ABB RAPID module: MAIN_1.prg

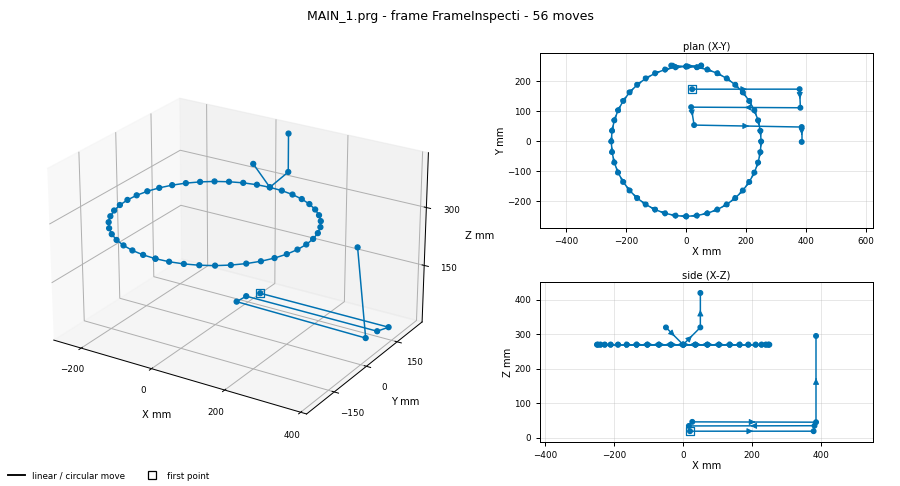
[picture p0: tool path of MAIN_1.prg in frame FrameInspecti, 56 of 76 moves have a stored position in this frame; points joined in program order, loops and branches not executed]
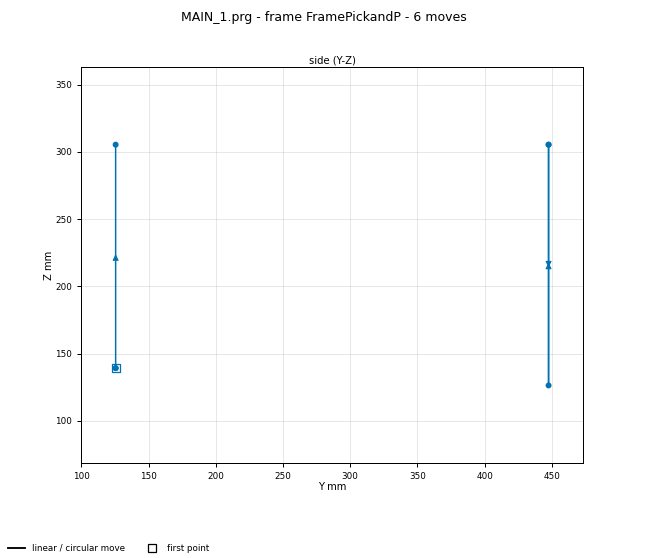
[picture p1: tool path of MAIN_1.prg in frame FramePickandP, 6 of 76 moves have a stored position in this frame; points joined in program order, loops and branches not executed]
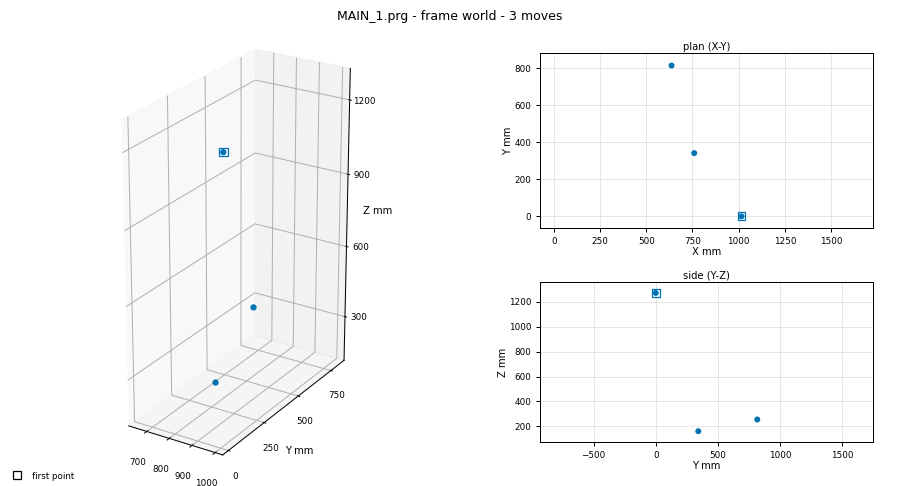
[picture p2: tool path of MAIN_1.prg in frame world, 3 of 76 moves have a stored position in this frame; points joined in program order, loops and branches not executed]
%%%
  VERSION:1
  LANGUAGE:ENGLISH
%%%
MODULE MOD_MAIN_1

    ! -------------------------------
    ! Define customized variables here
    ! ...

	! Tool variables:
	PERS tooldata Tool1 := [TRUE,[[129.073,0.000,85.477],[0.98018657,0.00000000,0.19807649,0.00000000]],[1,[0,0,20],[1,0,0,0],0,0,0.005]];
	PERS tooldata Tool1_withave := [TRUE,[[0.000,0.000,200.000],[1.00000000,0.00000000,0.00000000,0.00000000]],[1,[0,0,20],[1,0,0,0],0,0,0.005]];

	! Reference variables:
	PERS wobjdata FramePickandP := [FALSE, TRUE, "", [[719.013,-664.003,0.000],[1.00000000,0.00000000,0.00000000,0.00000000]],[[0,0,0],[1,0,0,0]]];
	PERS wobjdata FrameCircular := [FALSE, TRUE, "", [[577.670,392.250,0.000],[0.94275941,0.00000000,0.00000000,0.33347368]],[[0,0,0],[1,0,0,0]]];
	PERS wobjdata FrameInspecti := [FALSE, TRUE, "", [[0.000,782.714,377.610],[1.00000000,0.00000000,0.00000000,0.00000000]],[[0,0,0],[1,0,0,0]]];
	PERS wobjdata Frame1_withav := [FALSE, TRUE, "", [[0.000,1000.000,0.000],[1.00000000,0.00000000,0.00000000,0.00000000]],[[0,0,0],[1,0,0,0]]];

	PROC PROG1_withave()
		ConfJ \On;
		ConfL \Off;
		! This is a subprogram call to PROG_1
		MoveAbsJ [[-0.000001,0.000000,0.000000,0.000000,0.000000,-0.000000],[9E+09,9E+09,9E+09,9E+09,9E+09,9E+09]],v1000,z1,Tool1_withave \WObj:=Frame1_withav;
	ENDPROC

	PROC Main()
		ConfJ \On;
		ConfL \Off;
		! Program generated by RoboDK v5.6.9 for RoboDK Industrial on 26/02/2024 09:58:20
		! Using nominal kinematics.
		MoveAbsJ [[-0.000001,0.000000,0.000000,0.000000,0.000000,-0.000000],[9E+09,9E+09,9E+09,9E+09,9E+09,9E+09]],v500,z1,tool0 \WObj:=wobj0;
		MoveAbsJ [[0.000000,3.211240,-15.423700,0.000000,12.212500,-0.000000],[9E+09,9E+09,9E+09,9E+09,9E+09,9E+09]],v500,z1,tool0 \WObj:=wobj0;
		MoveL [[1015.000,0.000,1272.000],[0.70710678,0.00000000,0.70710678,0.00000001],[0,0,0,1],[9E+09,9E+09,9E+09,9E+09,9E+09,9E+09]],v500,z1,tool0 \WObj:=wobj0;
		SetDO D_OUT_5, 1;
		SetDO D_OUT_5, 1;
		SetDO D_OUT_5, 0.5;
		SetDO D_OUT_5, true;
		SetAO A_OUT_5, 1;
		SetAO A_OUT_5, 2;
		SetAO A_OUT_5, 0.5;
		SetAO A_OUT_5, true;
		SetDO var, val;
		SetAO var, val;
		WaitDI D_IN_5, 1;
		WaitDI D_IN_5, 1;
		WaitDI D_IN_5, 0.5;
		WaitDI D_IN_5, true;
		WaitDI D_IN_5, 1, \MaxTime:=0.1;
		WaitDI var, val;
		WaitDI var, val, \MaxTime:=0.1;
		TPWrite "Message";
		REMOTE_PROG_CALL_171;
		CODE_INSERT_172
		! Insert Comment
		MoveAbsJ [[-29.332200,46.677000,-0.024523,26.545600,25.395700,-51.634000],[9E+09,9E+09,9E+09,9E+09,9E+09,9E+09]],v500,z10,Tool1 \WObj:=FramePickandP;
		MoveL [[187.786,125.499,139.112],[0.00157079,-0.00002623,0.99999877,0.00003495],[-1,0,-1,0],[9E+09,9E+09,9E+09,9E+09,9E+09,9E+09]],v100,fine,Tool1 \WObj:=FramePickandP;
		SetDO D_OUT_5, 1;
		PICK_PART_111;
		MoveL CalcRobT([[-29.332200,46.677000,-0.024486,26.545800,25.395700,-51.634200],[9E+09,9E+09,9E+09,9E+09,9E+09,9E+09]],Tool1 \WObj:=FramePickandP),v300,z10,Tool1 \WObj:=FramePickandP;
		MoveL [[187.272,447.522,305.347],[0.00161443,0.00000875,0.99999870,-0.00001747],[-1,0,-1,0],[9E+09,9E+09,9E+09,9E+09,9E+09,9E+09]],v300,z10,Tool1 \WObj:=FramePickandP;
		! MoveSearch command not implemented
		MoveL [[187.851,447.517,126.235],[0.00161443,0.00000875,0.99999870,-0.00001747],[-1,0,-1,0],[9E+09,9E+09,9E+09,9E+09,9E+09,9E+09]],v100,fine,Tool1 \WObj:=FramePickandP;
		SetDO D_OUT_5, 0;
		PLACE_PART_112;
		MoveL [[187.272,447.522,305.347],[0.00161443,0.00000875,0.99999870,-0.00001747],[-1,0,-1,0],[9E+09,9E+09,9E+09,9E+09,9E+09,9E+09]],v100,z10,Tool1 \WObj:=FramePickandP;
		MoveAbsJ [[52.186000,45.675800,6.920000,66.734200,19.932300,-92.730000],[9E+09,9E+09,9E+09,9E+09,9E+09,9E+09]],v100,[FALSE,25.0,37.5,37.5,3.8,37.5,3.8],Tool1 \WObj:=FrameCircular;
		MoveC [[430.047,43.774,231.503],[0.08620627,-0.38531406,0.91758054,0.04634115],[0,0,-2,0],[9E+09,9E+09,9E+09,9E+09,9E+09,9E+09]],[[109.688,-153.222,161.073],[0.08620627,-0.38531406,0.91758054,0.04634115],[0,0,-2,0],[9E+09,9E+09,9E+09,9E+09,9E+09,9E+09]],v100,[FALSE,25.0,37.5,37.5,3.8,37.5,3.8],Tool1 \WObj:=FrameCircular;
		MoveC CalcRobT([[38.508400,52.810400,-4.822350,56.452300,29.788200,-93.025700],[9E+09,9E+09,9E+09,9E+09,9E+09,9E+09]], Tool1 \WObj:=FrameCircular),CalcRobT([[52.185900,45.675700,6.920040,66.734400,19.932300,-92.730300],[9E+09,9E+09,9E+09,9E+09,9E+09,9E+09]],Tool1 \WObj:=FrameCircular),v100,[FALSE,25.0,37.5,37.5,3.8,37.5,3.8],Tool1 \WObj:=FrameCircular;
		MoveL [[312.208,292.214,255.156],[0.08620627,-0.38531406,0.91758054,0.04634115],[0,0,-2,0],[9E+09,9E+09,9E+09,9E+09,9E+09,9E+09]],v100,fine,Tool1 \WObj:=FrameCircular;
		MoveAbsJ [[-0.000001,0.000000,0.000000,0.000000,0.000000,-0.000000],[9E+09,9E+09,9E+09,9E+09,9E+09,9E+09]],v100,fine,Tool1 \WObj:=FrameCircular;
		MoveAbsJ [[88.676000,29.601600,-6.428830,-1.984220,49.479200,4.547690],[9E+09,9E+09,9E+09,9E+09,9E+09,9E+09]],v100,fine,Tool1 \WObj:=FrameInspecti;
		MoveL [[19.898,174.307,19.008],[0.03212514,0.67543146,-0.73589088,0.03499889],[0,-1,0,0],[9E+09,9E+09,9E+09,9E+09,9E+09,9E+09]],v100,fine,Tool1 \WObj:=FrameInspecti;
		MoveL [[378.402,174.416,18.997],[0.03212514,0.67543146,-0.73589088,0.03499889],[0,0,-1,0],[9E+09,9E+09,9E+09,9E+09,9E+09,9E+09]],v100,fine,Tool1 \WObj:=FrameInspecti;
		MoveL [[380.996,112.363,34.882],[0.10687212,0.66688803,-0.72816340,0.11669088],[0,-1,-1,0],[9E+09,9E+09,9E+09,9E+09,9E+09,9E+09]],v100,fine,Tool1 \WObj:=FrameInspecti;
		MoveL [[16.551,114.359,34.226],[0.10687212,0.66688803,-0.72816340,0.11669088],[0,-1,0,0],[9E+09,9E+09,9E+09,9E+09,9E+09,9E+09]],v100,fine,Tool1 \WObj:=FrameInspecti;
		MoveL [[26.434,54.524,46.072],[0.02563823,-0.67223306,0.73935814,0.02819468],[0,-1,0,0],[9E+09,9E+09,9E+09,9E+09,9E+09,9E+09]],v100,fine,Tool1 \WObj:=FrameInspecti;
		MoveL [[385.448,48.050,45.137],[0.06581621,-0.66924184,0.73657112,0.07243323],[0,0,-1,0],[9E+09,9E+09,9E+09,9E+09,9E+09,9E+09]],v100,fine,Tool1 \WObj:=FrameInspecti;
		MoveL [[385.448,-1.625,295.251],[0.06581621,-0.66924184,0.73657112,0.07243323],[0,0,-1,0],[9E+09,9E+09,9E+09,9E+09,9E+09,9E+09]],v100,fine,Tool1 \WObj:=FrameInspecti;
		MoveAbsJ [[-0.000001,0.000000,0.000000,0.000000,0.000000,-0.000000],[9E+09,9E+09,9E+09,9E+09,9E+09,9E+09]],v100,fine,Tool1 \WObj:=FrameInspecti;
		EVENT_PROG_START_101;
		FrameInspecti := [FALSE, TRUE, "", [[13.637,-840.080,0.000],[0.70710678,0.00000000,0.00000000,-0.70710678]],[[0,0,0],[1,0,0,0]]];
		! Show Tool 1
		MoveAbsJ [[-68.090300,24.201900,26.785500,38.213400,36.201700,-98.796400],[9E+09,9E+09,9E+09,9E+09,9E+09,9E+09]],v1000,z1,Tool1 \WObj:=FrameInspecti;
		EVENT_PATH_APPROACH_102;
		MoveL [[-49.895,253.259,319.999],[0.00233251,-0.70710293,0.70710388,0.00202398],[-1,0,-2,0],[9E+09,9E+09,9E+09,9E+09,9E+09,9E+09]],v1000,z1,Tool1 \WObj:=FrameInspecti;
		MoveL [[0.000,250.000,270.000],[0.00233251,-0.70710293,0.70710388,0.00202398],[-1,0,-2,0],[9E+09,9E+09,9E+09,9E+09,9E+09,9E+09]],v1000,z1,Tool1 \WObj:=FrameInspecti;
		EVENT_PATH_START_103;
		MoveL [[35.579,247.455,270.000],[0.00259168,-0.70710203,0.70710482,0.00166608],[-1,0,-2,0],[9E+09,9E+09,9E+09,9E+09,9E+09,9E+09]],v50,z1,Tool1 \WObj:=FrameInspecti;
		MoveL [[70.433,239.873,270.000],[0.00280762,-0.70710738,0.70709946,0.00127734],[-1,0,-2,0],[9E+09,9E+09,9E+09,9E+09,9E+09,9E+09]],v50,z1,Tool1 \WObj:=FrameInspecti;
		MoveL [[103.854,227.408,270.000],[0.00295572,-0.70710677,0.70710008,0.00087007],[-1,0,-2,0],[9E+09,9E+09,9E+09,9E+09,9E+09,9E+09]],v50,z1,Tool1 \WObj:=FrameInspecti;
		MoveL [[135.160,210.313,270.000],[0.00305444,-0.70710635,0.70710047,0.00043812],[-1,0,-2,0],[9E+09,9E+09,9E+09,9E+09,9E+09,9E+09]],v50,z1,Tool1 \WObj:=FrameInspecti;
		MoveL [[163.715,188.937,270.000],[0.00308530,-0.70710622,0.70710061,0.00000001],[-1,0,-2,0],[9E+09,9E+09,9E+09,9E+09,9E+09,9E+09]],v50,z1,Tool1 \WObj:=FrameInspecti;
		MoveL [[188.937,163.715,270.000],[0.00305445,-0.70710635,0.70710047,-0.00043812],[-1,0,-2,0],[9E+09,9E+09,9E+09,9E+09,9E+09,9E+09]],v50,z1,Tool1 \WObj:=FrameInspecti;
		MoveL [[210.313,135.160,270.000],[0.00296806,-0.70710672,0.70710008,-0.00087007],[-1,0,-2,0],[9E+09,9E+09,9E+09,9E+09,9E+09,9E+09]],v50,z1,Tool1 \WObj:=FrameInspecti;
		MoveL [[227.408,103.854,270.000],[0.00281379,-0.70710735,0.70709945,-0.00128351],[-1,0,-2,0],[9E+09,9E+09,9E+09,9E+09,9E+09,9E+09]],v50,z1,Tool1 \WObj:=FrameInspecti;
		MoveL [[239.873,70.433,270.000],[0.00259785,-0.70710201,0.70710480,-0.00167225],[-1,0,-2,0],[9E+09,9E+09,9E+09,9E+09,9E+09,9E+09]],v50,z1,Tool1 \WObj:=FrameInspecti;
		MoveL [[247.455,35.579,270.000],[0.00233251,-0.70710293,0.70710388,-0.00202398],[-1,0,-2,0],[9E+09,9E+09,9E+09,9E+09,9E+09,9E+09]],v50,z1,Tool1 \WObj:=FrameInspecti;
		MoveL [[250.000,0.000,270.000],[0.00202398,-0.70710388,0.70710293,-0.00233251],[-1,0,-2,0],[9E+09,9E+09,9E+09,9E+09,9E+09,9E+09]],v50,z1,Tool1 \WObj:=FrameInspecti;
		MoveL [[247.455,-35.579,270.000],[0.00167225,-0.70710480,0.70710201,-0.00259785],[-1,0,-2,0],[9E+09,9E+09,9E+09,9E+09,9E+09,9E+09]],v50,z1,Tool1 \WObj:=FrameInspecti;
		MoveL [[239.873,-70.433,270.000],[0.00128351,-0.70709945,0.70710735,-0.00281379],[-2,0,-2,0],[9E+09,9E+09,9E+09,9E+09,9E+09,9E+09]],v50,z1,Tool1 \WObj:=FrameInspecti;
		MoveL [[227.408,-103.854,270.000],[0.00087007,-0.70710008,0.70710672,-0.00296806],[-2,0,-2,0],[9E+09,9E+09,9E+09,9E+09,9E+09,9E+09]],v50,z1,Tool1 \WObj:=FrameInspecti;
		MoveL [[210.313,-135.160,270.000],[0.00043812,-0.70710047,0.70710635,-0.00305445],[-2,0,-2,0],[9E+09,9E+09,9E+09,9E+09,9E+09,9E+09]],v50,z1,Tool1 \WObj:=FrameInspecti;
		MoveL [[188.937,-163.715,270.000],[0.00000000,-0.70710061,0.70710622,-0.00308530],[-2,0,-2,0],[9E+09,9E+09,9E+09,9E+09,9E+09,9E+09]],v50,z1,Tool1 \WObj:=FrameInspecti;
		MoveL [[163.715,-188.937,270.000],[0.00043812,0.70710047,-0.70710635,0.00305444],[-2,0,-2,0],[9E+09,9E+09,9E+09,9E+09,9E+09,9E+09]],v50,z1,Tool1 \WObj:=FrameInspecti;
		MoveL [[135.160,-210.313,270.000],[0.00087007,0.70710008,-0.70710672,0.00296806],[-2,0,-2,0],[9E+09,9E+09,9E+09,9E+09,9E+09,9E+09]],v50,z1,Tool1 \WObj:=FrameInspecti;
		MoveL [[103.854,-227.408,270.000],[0.00128351,0.70709945,-0.70710735,0.00281379],[-2,0,-2,0],[9E+09,9E+09,9E+09,9E+09,9E+09,9E+09]],v50,z1,Tool1 \WObj:=FrameInspecti;
		MoveL [[70.433,-239.873,270.000],[0.00167225,0.70710480,-0.70710201,0.00259785],[-2,0,-2,0],[9E+09,9E+09,9E+09,9E+09,9E+09,9E+09]],v50,z1,Tool1 \WObj:=FrameInspecti;
		MoveL [[35.579,-247.455,270.000],[0.00202398,0.70710388,-0.70710293,0.00233251],[-2,0,-2,0],[9E+09,9E+09,9E+09,9E+09,9E+09,9E+09]],v50,z1,Tool1 \WObj:=FrameInspecti;
		MoveL [[0.000,-250.000,270.000],[0.00202398,0.70710388,-0.70710293,0.00233251],[-2,0,-2,0],[9E+09,9E+09,9E+09,9E+09,9E+09,9E+09]],v50,z1,Tool1 \WObj:=FrameInspecti;
		MoveL [[0.000,-250.000,270.000],[0.00233251,0.70710293,-0.70710388,0.00202398],[-2,0,-2,0],[9E+09,9E+09,9E+09,9E+09,9E+09,9E+09]],v50,z1,Tool1 \WObj:=FrameInspecti;
		MoveL [[-35.579,-247.455,270.000],[0.00259785,0.70710201,-0.70710480,0.00167225],[-2,0,-2,0],[9E+09,9E+09,9E+09,9E+09,9E+09,9E+09]],v50,z1,Tool1 \WObj:=FrameInspecti;
		MoveL [[-70.433,-239.873,270.000],[0.00280762,0.70710738,-0.70709946,0.00127734],[-2,0,-2,0],[9E+09,9E+09,9E+09,9E+09,9E+09,9E+09]],v50,z1,Tool1 \WObj:=FrameInspecti;
		MoveL [[-103.854,-227.408,270.000],[0.00295572,0.70710677,-0.70710008,0.00087007],[-2,0,-2,0],[9E+09,9E+09,9E+09,9E+09,9E+09,9E+09]],v50,z1,Tool1 \WObj:=FrameInspecti;
		MoveL [[-135.160,-210.313,270.000],[0.00305444,0.70710635,-0.70710047,0.00043812],[-2,0,-2,0],[9E+09,9E+09,9E+09,9E+09,9E+09,9E+09]],v50,z1,Tool1 \WObj:=FrameInspecti;
		MoveL [[-163.715,-188.937,270.000],[0.00308530,0.70710622,-0.70710061,0.00000001],[-2,0,-2,0],[9E+09,9E+09,9E+09,9E+09,9E+09,9E+09]],v50,z1,Tool1 \WObj:=FrameInspecti;
		MoveL [[-188.937,-163.715,270.000],[0.00305445,0.70710635,-0.70710047,-0.00043812],[-2,0,-2,0],[9E+09,9E+09,9E+09,9E+09,9E+09,9E+09]],v50,z1,Tool1 \WObj:=FrameInspecti;
		MoveL [[-210.313,-135.160,270.000],[0.00295572,0.70710677,-0.70710008,-0.00087007],[-2,0,-2,0],[9E+09,9E+09,9E+09,9E+09,9E+09,9E+09]],v50,z1,Tool1 \WObj:=FrameInspecti;
		MoveL [[-227.408,-103.854,270.000],[0.00280145,0.70710740,-0.70709945,-0.00128351],[-2,0,-2,0],[9E+09,9E+09,9E+09,9E+09,9E+09,9E+09]],v50,z1,Tool1 \WObj:=FrameInspecti;
		MoveL [[-239.873,-70.433,270.000],[0.00259785,0.70710201,-0.70710480,-0.00167225],[-2,0,-2,0],[9E+09,9E+09,9E+09,9E+09,9E+09,9E+09]],v50,z1,Tool1 \WObj:=FrameInspecti;
		MoveL [[-247.455,-35.579,270.000],[0.00233251,0.70710293,-0.70710388,-0.00202398],[-1,0,-2,0],[9E+09,9E+09,9E+09,9E+09,9E+09,9E+09]],v50,z1,Tool1 \WObj:=FrameInspecti;
		MoveL [[-250.000,0.000,270.000],[0.00202398,0.70710388,-0.70710293,-0.00233251],[-1,0,-2,0],[9E+09,9E+09,9E+09,9E+09,9E+09,9E+09]],v50,z1,Tool1 \WObj:=FrameInspecti;
		MoveL [[-247.455,35.579,270.000],[0.00166608,0.70710482,-0.70710203,-0.00259168],[-1,0,-2,0],[9E+09,9E+09,9E+09,9E+09,9E+09,9E+09]],v50,z1,Tool1 \WObj:=FrameInspecti;
		MoveL [[-239.873,70.433,270.000],[0.00128351,0.70709945,-0.70710740,-0.00280145],[-1,0,-2,0],[9E+09,9E+09,9E+09,9E+09,9E+09,9E+09]],v50,z1,Tool1 \WObj:=FrameInspecti;
		MoveL [[-227.408,103.854,270.000],[0.00087007,0.70710008,-0.70710672,-0.00296806],[-1,0,-2,0],[9E+09,9E+09,9E+09,9E+09,9E+09,9E+09]],v50,z1,Tool1 \WObj:=FrameInspecti;
		MoveL [[-210.313,135.160,270.000],[0.00043812,0.70710047,-0.70710635,-0.00305445],[-1,0,-2,0],[9E+09,9E+09,9E+09,9E+09,9E+09,9E+09]],v50,z1,Tool1 \WObj:=FrameInspecti;
		MoveL [[-188.937,163.715,270.000],[0.00000000,-0.70710061,0.70710622,0.00308530],[-1,0,-2,0],[9E+09,9E+09,9E+09,9E+09,9E+09,9E+09]],v50,z1,Tool1 \WObj:=FrameInspecti;
		MoveL [[-163.715,188.937,270.000],[0.00043812,-0.70710047,0.70710635,0.00305444],[-1,0,-2,0],[9E+09,9E+09,9E+09,9E+09,9E+09,9E+09]],v50,z1,Tool1 \WObj:=FrameInspecti;
		MoveL [[-135.160,210.313,270.000],[0.00087007,-0.70710008,0.70710677,0.00295572],[-1,0,-2,0],[9E+09,9E+09,9E+09,9E+09,9E+09,9E+09]],v50,z1,Tool1 \WObj:=FrameInspecti;
		MoveL [[-103.854,227.408,270.000],[0.00128351,-0.70709945,0.70710735,0.00281379],[-1,0,-2,0],[9E+09,9E+09,9E+09,9E+09,9E+09,9E+09]],v50,z1,Tool1 \WObj:=FrameInspecti;
		MoveL [[-70.433,239.873,270.000],[0.00167225,-0.70710480,0.70710201,0.00259785],[-1,0,-2,0],[9E+09,9E+09,9E+09,9E+09,9E+09,9E+09]],v50,z1,Tool1 \WObj:=FrameInspecti;
		MoveL [[-35.579,247.455,270.000],[0.00202398,-0.70710388,0.70710293,0.00233251],[-1,0,-2,0],[9E+09,9E+09,9E+09,9E+09,9E+09,9E+09]],v50,z1,Tool1 \WObj:=FrameInspecti;
		MoveL [[0.000,250.000,270.000],[0.00202398,-0.70710388,0.70710293,0.00233251],[-1,0,-2,0],[9E+09,9E+09,9E+09,9E+09,9E+09,9E+09]],v50,z1,Tool1 \WObj:=FrameInspecti;
		EVENT_PATH_FINISH_105;
		MoveL [[49.895,253.258,319.999],[0.00202398,-0.70710388,0.70710293,0.00233251],[-1,0,-2,0],[9E+09,9E+09,9E+09,9E+09,9E+09,9E+09]],v1000,z1,Tool1 \WObj:=FrameInspecti;
		MoveL [[49.939,252.642,419.997],[0.00202398,-0.70710388,0.70710293,0.00233251],[-1,0,-2,0],[9E+09,9E+09,9E+09,9E+09,9E+09,9E+09]],v1000,z1,Tool1 \WObj:=FrameInspecti;
		EVENT_PATH_RETRACT_106;
		EVENT_PROG_FINISH_107;
		FramePickandP := [FALSE, TRUE, "", [[719.013,-664.003,0.000],[1.00000000,0.00000000,0.00000000,0.00000000]],[[0,0,0],[1,0,0,0]]];
		MoveAbsJ [[-29.332200,46.677000,-0.024523,26.545600,25.395700,-51.634000],[9E+09,9E+09,9E+09,9E+09,9E+09,9E+09]],v1000,z1,Tool1 \WObj:=FramePickandP;
		WaitTime 1.250;
		MoveL [[187.786,125.499,139.112],[0.00157079,-0.00002623,0.99999877,0.00003495],[-1,0,-1,0],[9E+09,9E+09,9E+09,9E+09,9E+09,9E+09]],v1000,z1,Tool1 \WObj:=FramePickandP;
		WaitDI D_IN_1, 1;
		MoveL [[187.264,125.487,305.356],[0.00160570,0.00000000,0.99999871,-0.00000000],[-1,0,-1,0],[9E+09,9E+09,9E+09,9E+09,9E+09,9E+09]],v1000,z1,Tool1 \WObj:=FramePickandP;
		PROG1_withaverylongnameandspecialcharacters;
	ENDPROC

ENDMODULE
